(* IEC 61131-3 sources: sis-interlock-demo/src/POUs/Sis/F_CemCheckCfg, 2 files *)

(* ---- F_CemCheckCfg.decl.st ---- *)
// Назначение: проверка конфигурации матрицы: сумма битов CEM_CFG_* (таблица 4.3); 0 — верна.
//             При CEM_CFG_COUNT причины и следствия не проверяются, CRC проверяется всегда.
//             Используемая причина — i <= uiCauseCount (включена она или нет), используемое
//             следствие — j <= uiEffectCount. Разрешённый обход: срок в (0, SIS_OVERRIDE_MAX],
//             подтверждение нормы для автоснятия в (0, tOverrideMax).
// Автор:      kr0nsch
// Версия:     0.2.0
// Документ:   docs/DESIGN.md, раздел «6.8 Конфигурация и CRC»
// ВНИМАНИЕ:   код демонстрационный и не предназначен для систем безопасности. Реальная ПАЗ
//             требует определения SIL, сертифицированных аппаратных и программных средств
//             и валидации по ГОСТ Р МЭК 61511.
FUNCTION F_CemCheckCfg : WORD
VAR_IN_OUT CONSTANT
    stCfg : ST_CemCfg;   // проверяемая конфигурация
END_VAR
VAR
    wErr       : WORD;          // найденные ошибки
    wUsedMask  : WORD;          // биты используемых причин
    uiI        : UINT;          // индекс причины
    uiJ        : UINT;          // индекс следствия
    stCause    : ST_CauseCfg;   // копия строки
    stEffect   : ST_EffectCfg;  // копия столбца
    xSourceOk  : BOOL;          // источник требования из перечисления
    xOvrTimeOk : BOOL;          // длительность обхода в (0, SIS_OVERRIDE_MAX]
    xOvrClrOk  : BOOL;          // подтверждение нормы для автоснятия обхода в (0, tOverrideMax)
    xSafeOk    : BOOL;          // безопасное состояние из перечисления
    xCauseBad  : BOOL;          // есть неверная причина
    xEffectBad : BOOL;          // есть неверное следствие
END_VAR

(* ---- F_CemCheckCfg.impl.st ---- *)
wErr := 0;
xCauseBad := FALSE;
xEffectBad := FALSE;

IF stCfg.uiCauseCount < 1 OR stCfg.uiCauseCount > GVL_Const.SIS_CAUSES_MAX
    OR stCfg.uiEffectCount < 1 OR stCfg.uiEffectCount > GVL_Const.SIS_EFFECTS_MAX
THEN
    wErr := wErr OR GVL_Const.CEM_CFG_COUNT;
ELSE
    // Причины: источник, предел задержки, срок разрешённого обхода и подтверждение нормы для его
    // автоснятия — короче срока, иначе обход не снимется при норме раньше срока (6.4)
    FOR uiI := 1 TO stCfg.uiCauseCount DO
        stCause := stCfg.astCause[uiI];
        xSourceOk := stCause.eSource = E_CauseSource.Voting OR stCause.eSource = E_CauseSource.External;
        xOvrTimeOk := stCause.tOverrideMax > T#0S AND stCause.tOverrideMax <= GVL_Const.SIS_OVERRIDE_MAX;
        xOvrClrOk := stCause.tOverrideClear > T#0S AND stCause.tOverrideClear < stCause.tOverrideMax;
        IF NOT xSourceOk OR stCause.tDelay > GVL_Const.SIS_DELAY_MAX
            OR (stCause.xOverrideAllowed AND NOT (xOvrTimeOk AND xOvrClrOk))
        THEN
            xCauseBad := TRUE;
        END_IF
    END_FOR

    // Следствия: используемые — состояние из перечисления, маска не пуста и без причин сверх
    // uiCauseCount; неиспользуемые — пустая маска
    wUsedMask := F_SisLowMask(uiCount := stCfg.uiCauseCount);
    FOR uiJ := 1 TO GVL_Const.SIS_EFFECTS_MAX DO
        stEffect := stCfg.astEffect[uiJ];
        IF uiJ <= stCfg.uiEffectCount THEN
            xSafeOk := stEffect.eSafeState = E_SafeState.Closed OR stEffect.eSafeState = E_SafeState.Open
                OR stEffect.eSafeState = E_SafeState.Stopped OR stEffect.eSafeState = E_SafeState.Off
                OR stEffect.eSafeState = E_SafeState.Alarm;
            IF NOT xSafeOk OR stEffect.wCauseMask = 0 OR (stEffect.wCauseMask AND NOT wUsedMask) <> 0 THEN
                xEffectBad := TRUE;
            END_IF
        ELSIF stEffect.wCauseMask <> 0 THEN
            xEffectBad := TRUE;
        END_IF
    END_FOR

    IF xCauseBad THEN
        wErr := wErr OR GVL_Const.CEM_CFG_CAUSE;
    END_IF
    IF xEffectBad THEN
        wErr := wErr OR GVL_Const.CEM_CFG_EFFECT;
    END_IF
END_IF

// CRC — всегда
IF F_CemCrc(stCfg := stCfg) <> stCfg.wMatrixCrc THEN
    wErr := wErr OR GVL_Const.CEM_CFG_CRC;
END_IF

F_CemCheckCfg := wErr;
